FUNCTION_BLOCK FB_ErrorCollector
VAR_INPUT
END_VAR
VAR_OUTPUT
END_VAR
VAR
	i: INT;
END_VAR

METHOD M_NewError : BOOL
VAR_INPUT
	eID:	E_ErrorIDs;
	eSrc:	E_ErrorSrcs;
	sMsg: 	STRING;
END_VAR
FOR i := 0 TO HMI.nNumberErrors - 1 DO
	IF HMI.aErrors[i].nType = eID AND HMI.aErrors[i].nSource = eSrc THEN
		RETURN;
	END_IF
END_FOR

HMI.aErrors[HMI.nNumberErrors].nType := eID;
HMI.aErrors[HMI.nNumberErrors].nSource := eSrc;
HMI.aErrors[HMI.nNumberErrors].sMsg := sMsg;
HMI.nNumberErrors := HMI.nNumberErrors + 1;
HMI.bErrorChange := TRUE;
END_METHOD

METHOD M_QuitError : BOOL
VAR_INPUT
	eID:	E_ErrorIDs;
	eSrc:	E_ErrorSrcs;
END_VAR
FOR i := 0 TO HMI.nNumberErrors - 1 DO
	IF HMI.aErrors[i].nType = eID AND HMI.aErrors[i].nSource = eSrc THEN
		MEMSET(ADR(HMI.aErrors[i]), 0, SIZEOF(HMI.aErrors[i]));
		IF NOT (i = MAX_ERRORS - 1) THEN
			MEMMOVE(ADR(HMI.aErrors[i]), ADR(HMI.aErrors[i + 1]), SIZEOF(HMI.aErrors[i]) * HMI.nNumberErrors - i - 1);
			MEMSET(ADR(HMI.aErrors[HMI.nNumberErrors - 1]), 0, SIZEOF(HMI.aErrors[HMI.nNumberErrors - 1]));
		END_IF
		HMI.nNumberErrors := HMI.nNumberErrors - 1;
		HMI.bErrorChange := TRUE;
		EXIT;
	END_IF
END_FOR
END_METHOD

END_FUNCTION_BLOCK

(* stored: Version 1.1.0.1, ProductVersion 3.1.4024.12
   POU FB_ErrorCollector: Id {f9aa26c4-0483-423f-82a5-7b8beceaf572}, SpecialFunc None
   Method M_NewError: Id {924919ae-eecd-4203-ba52-ec4cc691f278}
   Method M_QuitError: Id {7ec86467-9e08-471d-b1ed-7c539d76da3c} *)
